FUNCTION_BLOCK ABSTRACT FB_LogRecordProcessor_Base

METHOD ABSTRACT enrich
VAR_IN_OUT
	logRecord: FB_LogRecord;
END_VAR
END_METHOD

METHOD ABSTRACT free
VAR_INPUT
END_VAR
END_METHOD

METHOD ABSTRACT onEmit
VAR_INPUT
	logRecord: REFERENCE TO FB_LogRecord;
END_VAR
END_METHOD

PROPERTY pSelf : POINTER TO FB_LogRecordProcessor_Base
GET
pSelf := THIS;
END_GET
END_PROPERTY

METHOD ABSTRACT tick
END_METHOD

END_FUNCTION_BLOCK

(* stored: Version 1.1.0.1
   POU FB_LogRecordProcessor_Base: Id {aa1bfa7c-b5dc-4612-a924-12e642b6c02f}, SpecialFunc None
   Method enrich: Id {3eac3c59-065f-4409-b093-3f236ed38136}
   Method free: Id {bb9a97e7-e8b6-435b-b60a-d9e1aed96714}
   Method onEmit: Id {78085cb7-8a8c-4a0b-944f-aabfe8e6f9b1}
   Property pSelf: Id {0cb5a61d-3f85-49f6-b36f-cbe42579cdfb}
   Get Get: Id {992ce7aa-726b-498b-82b0-d35f11b9aaaa}
   Method tick: Id {63f82bb7-f9fd-41ad-8b62-442fb408f861} *)
